(* Logix 5000 project; controller NWGG 1756-L72 rev 35.12; software revision 35.00; part 18 of 19 *)
(* tags used below, declared in another part *)
   Auto_Start_Treatment : BOOL;
   Belt : udt_Motor[16];
   Belts_Ready : BOOL;
   Bin_Gate_Test : BOOL;
   Bin_Open_test : BOOL;
   Bins_Rqd : BOOL;
   ckIDX : DINT;
   cntTransferTime : COUNTER;
   cntTreatTime : COUNTER;
   Concrete_Belts_Ready : BOOL;
   Concrete_Leg : udt_Motor;
   Current_Dist_List_IDX : DINT;
   Finish_Treat_Ok : BOOL;
   IDX : DINT;
   Loadout_Bin : udt_Loadout_Bin[29];
   Loadout_K_Valve : udt_Loadout_K_Valve[2];
   Longest_Treat_Stop_IDX : DINT;
   Loop_Idx : DINT;
   Manual_Mode : BOOL;
   Pause_Load_By_Time : BOOL[32];
   Pause_Load_By_Weight : BOOL[32];
   Pause_Load_Expired : DINT[2];
   Pause_Load_Pre : DINT[2];
   Pause_Transfer_By_Time : BOOL;
   Pause_Transfer_Load_Expired : DINT;
   Pause_Transfer_Msc : DINT;
   Pause_Transfer_Pre : DINT;
   Remote_Pause_Treat : BOOL;
   Reset_Remote_Pause : BOOL;
   Reset_Treat_Chemicals : BOOL;
   Reversing_Belt_Bypass_Valve : BOOL;
   Reversing_Belt_Reversed : BOOL;
   Start_Treat_Belts_Enabled : BOOL;
   Steel_Rqd_Belts_Running : BOOL;
   Stop_Treater : BOOL;
   Target_Weight : DINT[2];
   tmr_Pause_Load_Timer : TIMER[2];
   tmr_Pause_Transfer_Timer : TIMER;
   tmrBin_Delay_Start : TIMER[30];
   tmrDelayTreatStart : TIMER;
   tmrDelayTreatStop : TIMER;
   tmrResetChemicals : TIMER;
   tmrTransferTime : TIMER;
   tmrTreatTime : TIMER;
   Transfer_Batch_Status : DINT;
   Transfer_Belts_Starting : BOOL;
   Transfer_From_IDX : DINT;
   Transfer_Interlock : BOOL;
   Transfer_To_IDX : DINT;
   TransferHours : DINT;
   TransferMinuets : DINT;
   TransferSeconds : DINT;
   Treat_Batch_Status : DINT;
   Treat_Bin_Gates_Opened : BOOL;
   Treat_Bins_Open : BOOL;
   Treat_Interlock : BOOL;
   Treater_Loadout : udt_Treater_Loadout;
   TreatHours : DINT;
   Treatment_Running : BOOL;
   Treatment_Started : BOOL;
   TreatMinuets : DINT;
   TreatSeconds : DINT;
   Use_Concrete_Side_Treat : BOOL;
   Use_Steel_Side_Treat : BOOL;
   Use_Steel_Transfer_Bins : BOOL;
   tmrSetWaterOil : TIMER;
   Treater_Remote_Out : DINT;
   Truck_Scales : udt_Truck_Scale[2];
(* SeedLoadoutMain, continued *)

ROUTINE tmrTest   (* ladder *)
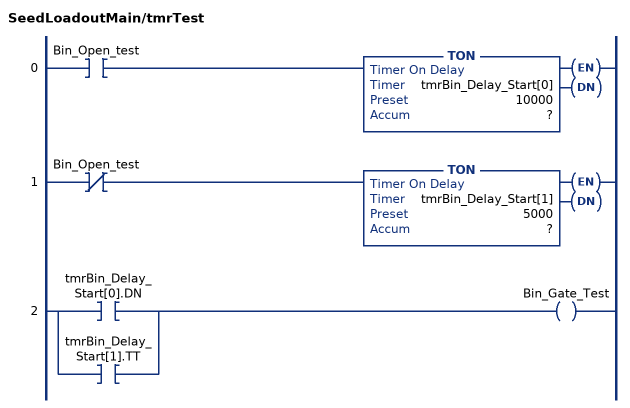
   0: XIC(Bin_Open_test)TON(tmrBin_Delay_Start[0],?,?);
   1: XIO(Bin_Open_test)TON(tmrBin_Delay_Start[1],?,?);
   2: [XIC(tmrBin_Delay_Start[0].DN) ,XIC(tmrBin_Delay_Start[1].TT) ]OTE(Bin_Gate_Test);
END_ROUTINE

ROUTINE Transfer_Belt_Batch_Ready   (* ladder *)
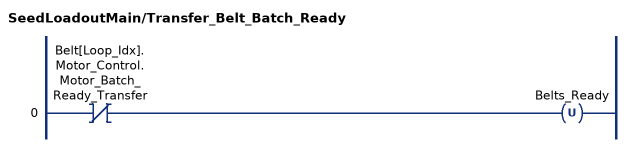
   0: XIO(Belt[Loop_Idx].Motor_Control.Motor_Batch_Ready_Transfer)OTU(Belts_Ready);
END_ROUTINE

ROUTINE Transfer_Belt_Start   (* ladder *)
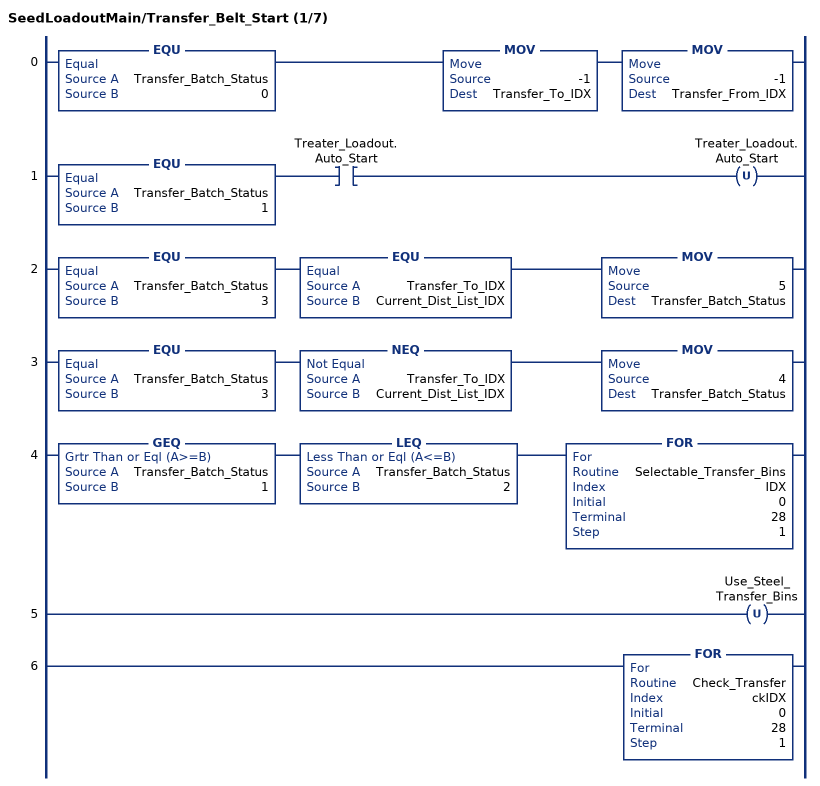
   0: EQU(Transfer_Batch_Status,0)MOV(-1,Transfer_To_IDX)MOV(-1,Transfer_From_IDX);
   1: EQU(Transfer_Batch_Status,1)XIC(Treater_Loadout.Auto_Start)OTU(Treater_Loadout.Auto_Start);
   2: EQU(Transfer_Batch_Status,3)EQU(Transfer_To_IDX,Current_Dist_List_IDX)MOV(5,Transfer_Batch_Status);
   3: EQU(Transfer_Batch_Status,3)NEQ(Transfer_To_IDX,Current_Dist_List_IDX)MOV(4,Transfer_Batch_Status);
   4: GEQ(Transfer_Batch_Status,1)LEQ(Transfer_Batch_Status,2)FOR(Selectable_Transfer_Bins,IDX,0,28,1);
   5: OTU(Use_Steel_Transfer_Bins);
   6: FOR(Check_Transfer,ckIDX,0,28,1);
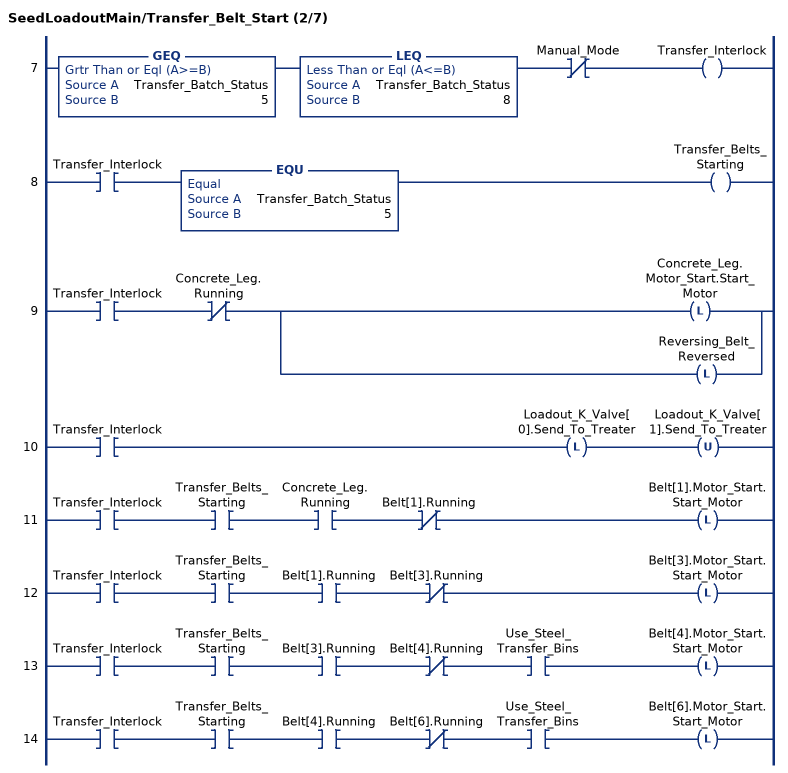
   7: GEQ(Transfer_Batch_Status,5)LEQ(Transfer_Batch_Status,8)XIO(Manual_Mode)OTE(Transfer_Interlock);
   8: XIC(Transfer_Interlock)EQU(Transfer_Batch_Status,5)OTE(Transfer_Belts_Starting);
   9: XIC(Transfer_Interlock)XIO(Concrete_Leg.Running)[OTL(Concrete_Leg.Motor_Start.Start_Motor) ,OTL(Reversing_Belt_Reversed) ];
   10: XIC(Transfer_Interlock)OTL(Loadout_K_Valve[0].Send_To_Treater)OTU(Loadout_K_Valve[1].Send_To_Treater);
   11: XIC(Transfer_Interlock)XIC(Transfer_Belts_Starting)XIC(Concrete_Leg.Running)XIO(Belt[1].Running)OTL(Belt[1].Motor_Start.Start_Motor);
   12: XIC(Transfer_Interlock)XIC(Transfer_Belts_Starting)XIC(Belt[1].Running)XIO(Belt[3].Running)OTL(Belt[3].Motor_Start.Start_Motor);
   13: XIC(Transfer_Interlock)XIC(Transfer_Belts_Starting)XIC(Belt[3].Running)XIO(Belt[4].Running)XIC(Use_Steel_Transfer_Bins)OTL(Belt[4].Motor_Start.Start_Motor);
   14: XIC(Transfer_Interlock)XIC(Transfer_Belts_Starting)XIC(Belt[4].Running)XIO(Belt[6].Running)XIC(Use_Steel_Transfer_Bins)OTL(Belt[6].Motor_Start.Start_Motor);
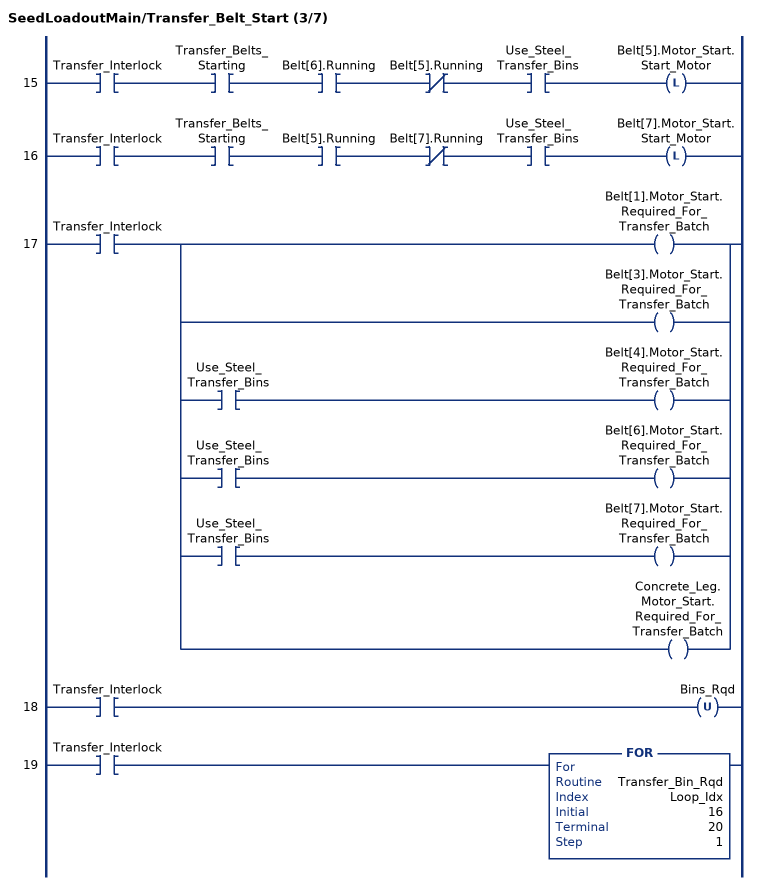
   15: XIC(Transfer_Interlock)XIC(Transfer_Belts_Starting)XIC(Belt[6].Running)XIO(Belt[5].Running)XIC(Use_Steel_Transfer_Bins)OTL(Belt[5].Motor_Start.Start_Motor);
   16: XIC(Transfer_Interlock)XIC(Transfer_Belts_Starting)XIC(Belt[5].Running)XIO(Belt[7].Running)XIC(Use_Steel_Transfer_Bins)OTL(Belt[7].Motor_Start.Start_Motor);
   17: XIC(Transfer_Interlock)[OTE(Belt[1].Motor_Start.Required_For_Transfer_Batch) ,OTE(Belt[3].Motor_Start.Required_For_Transfer_Batch) ,XIC(Use_Steel_Transfer_Bins) OTE(Belt[4].Motor_Start.Required_For_Transfer_Batch) ,XIC(Use_Steel_Transfer_Bins) OTE(Belt[6].Motor_Start.Required_For_Transfer_Batch) ,XIC(Use_Steel_Transfer_Bins) OTE(Belt[7].Motor_Start.Required_For_Transfer_Batch) ,OTE(Concrete_Leg.Motor_Start.Required_For_Transfer_Batch) ];
   18: XIC(Transfer_Interlock)OTU(Bins_Rqd);
   19: XIC(Transfer_Interlock)FOR(Transfer_Bin_Rqd,Loop_Idx,16,20,1);
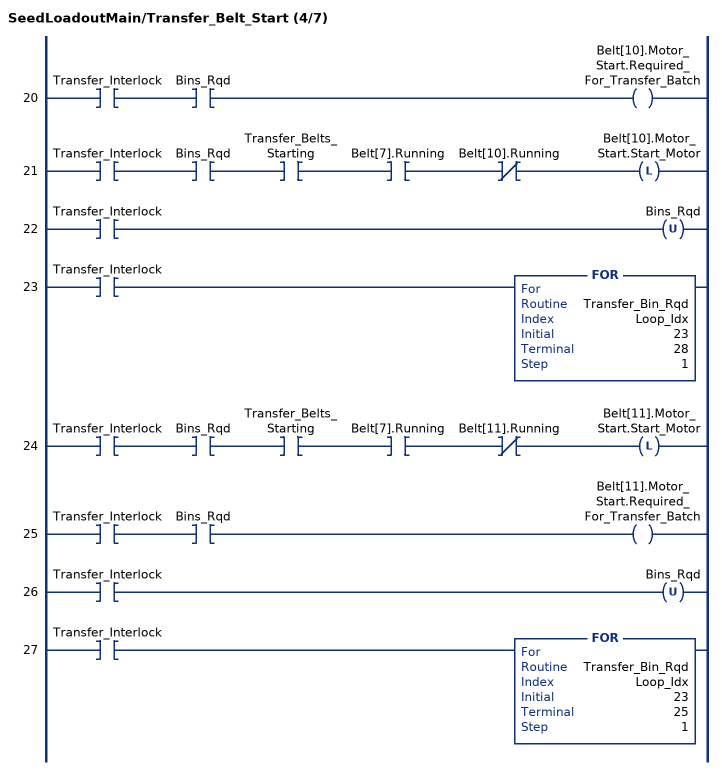
   20: XIC(Transfer_Interlock)XIC(Bins_Rqd)OTE(Belt[10].Motor_Start.Required_For_Transfer_Batch);
   21: XIC(Transfer_Interlock)XIC(Bins_Rqd)XIC(Transfer_Belts_Starting)XIC(Belt[7].Running)XIO(Belt[10].Running)OTL(Belt[10].Motor_Start.Start_Motor);
   22: XIC(Transfer_Interlock)OTU(Bins_Rqd);
   23: XIC(Transfer_Interlock)FOR(Transfer_Bin_Rqd,Loop_Idx,23,28,1);
   24: XIC(Transfer_Interlock)XIC(Bins_Rqd)XIC(Transfer_Belts_Starting)XIC(Belt[7].Running)XIO(Belt[11].Running)OTL(Belt[11].Motor_Start.Start_Motor);
   25: XIC(Transfer_Interlock)XIC(Bins_Rqd)OTE(Belt[11].Motor_Start.Required_For_Transfer_Batch);
   26: XIC(Transfer_Interlock)OTU(Bins_Rqd);
   27: XIC(Transfer_Interlock)FOR(Transfer_Bin_Rqd,Loop_Idx,23,25,1);
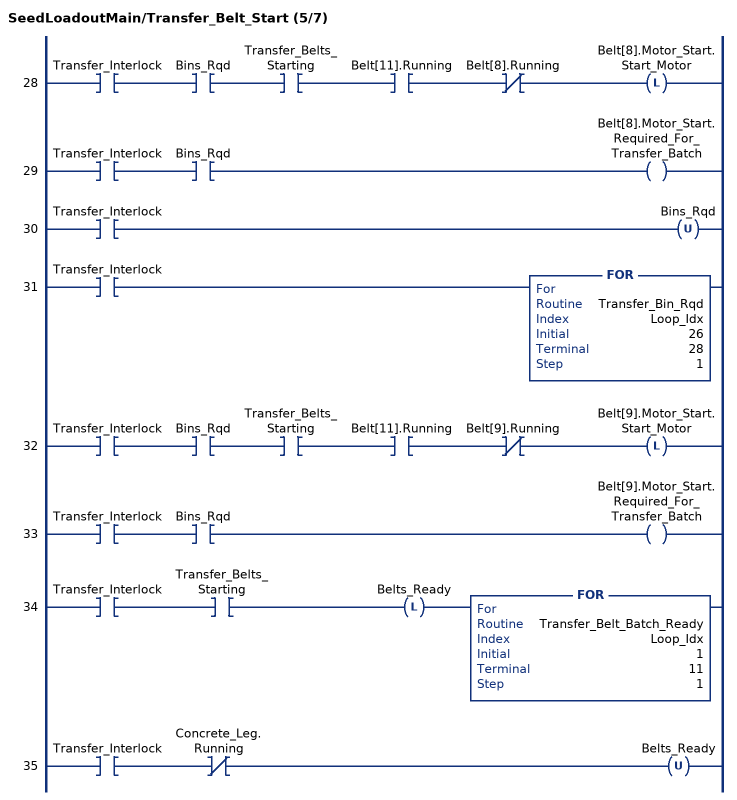
   28: XIC(Transfer_Interlock)XIC(Bins_Rqd)XIC(Transfer_Belts_Starting)XIC(Belt[11].Running)XIO(Belt[8].Running)OTL(Belt[8].Motor_Start.Start_Motor);
   29: XIC(Transfer_Interlock)XIC(Bins_Rqd)OTE(Belt[8].Motor_Start.Required_For_Transfer_Batch);
   30: XIC(Transfer_Interlock)OTU(Bins_Rqd);
   31: XIC(Transfer_Interlock)FOR(Transfer_Bin_Rqd,Loop_Idx,26,28,1);
   32: XIC(Transfer_Interlock)XIC(Bins_Rqd)XIC(Transfer_Belts_Starting)XIC(Belt[11].Running)XIO(Belt[9].Running)OTL(Belt[9].Motor_Start.Start_Motor);
   33: XIC(Transfer_Interlock)XIC(Bins_Rqd)OTE(Belt[9].Motor_Start.Required_For_Transfer_Batch);
   34: XIC(Transfer_Interlock)XIC(Transfer_Belts_Starting)OTL(Belts_Ready)FOR(Transfer_Belt_Batch_Ready,Loop_Idx,1,11,1);
   35: XIC(Transfer_Interlock)XIO(Concrete_Leg.Running)OTU(Belts_Ready);
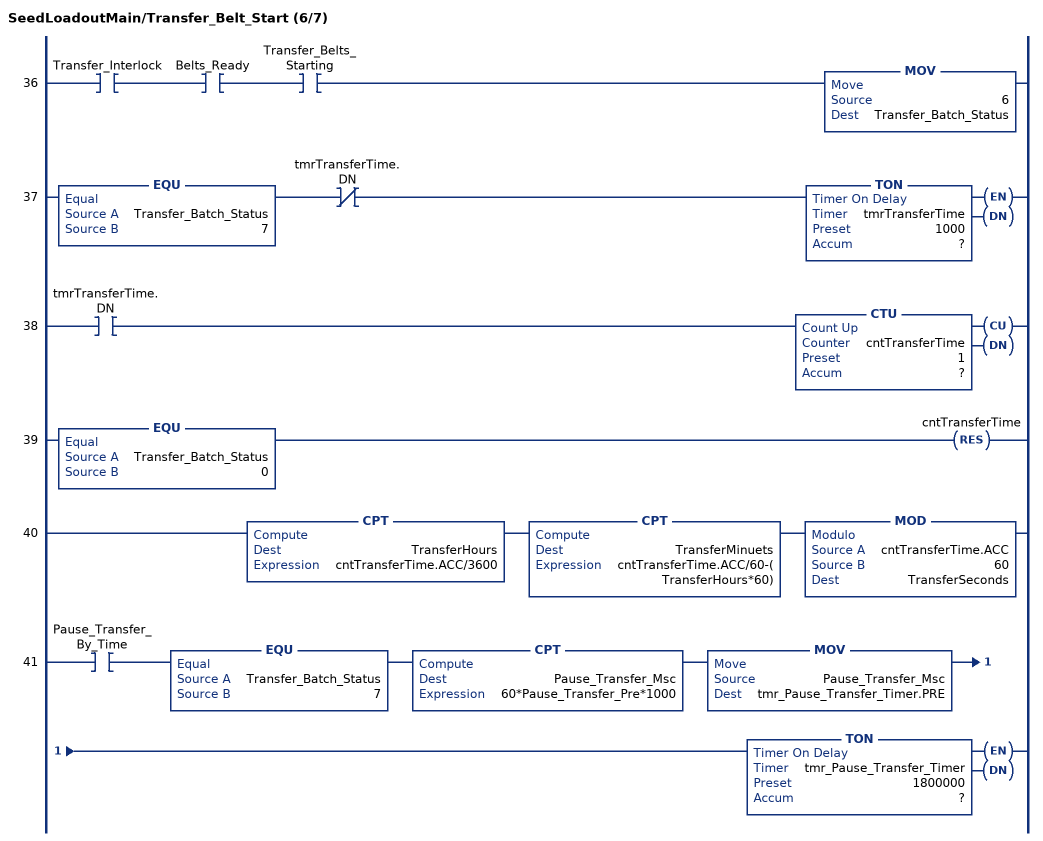
   36: XIC(Transfer_Interlock)XIC(Belts_Ready)XIC(Transfer_Belts_Starting)MOV(6,Transfer_Batch_Status);
   37: EQU(Transfer_Batch_Status,7)XIO(tmrTransferTime.DN)TON(tmrTransferTime,?,?);
   38: XIC(tmrTransferTime.DN)CTU(cntTransferTime,?,?);
   39: EQU(Transfer_Batch_Status,0)RES(cntTransferTime);
   40: CPT(TransferHours,cntTransferTime.ACC/3600)CPT(TransferMinuets,cntTransferTime.ACC/60-(TransferHours*60))MOD(cntTransferTime.ACC,60,TransferSeconds);
   41: XIC(Pause_Transfer_By_Time)EQU(Transfer_Batch_Status,7)CPT(Pause_Transfer_Msc,60*Pause_Transfer_Pre*1000)MOV(Pause_Transfer_Msc,tmr_Pause_Transfer_Timer.PRE)TON(tmr_Pause_Transfer_Timer,?,?);
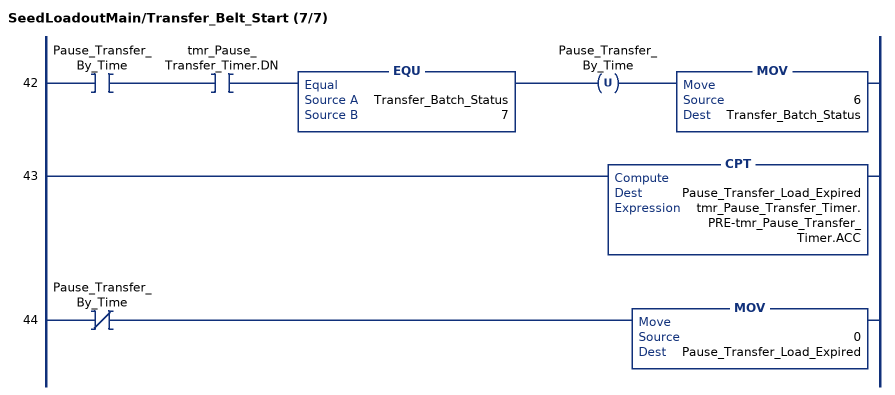
   42: XIC(Pause_Transfer_By_Time)XIC(tmr_Pause_Transfer_Timer.DN)EQU(Transfer_Batch_Status,7)OTU(Pause_Transfer_By_Time)MOV(6,Transfer_Batch_Status);
   43: CPT(Pause_Transfer_Load_Expired,tmr_Pause_Transfer_Timer.PRE-tmr_Pause_Transfer_Timer.ACC);
   44: XIO(Pause_Transfer_By_Time)MOV(0,Pause_Transfer_Load_Expired);
END_ROUTINE

ROUTINE Transfer_Bin_Rqd   (* ladder *)
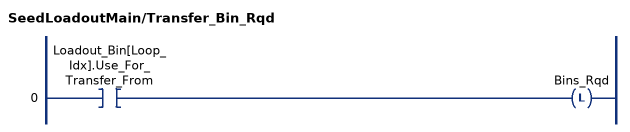
   0: XIC(Loadout_Bin[Loop_Idx].Use_For_Transfer_From)OTL(Bins_Rqd);
END_ROUTINE

ROUTINE Treat_Belt_Batch_Ready   (* ladder *)
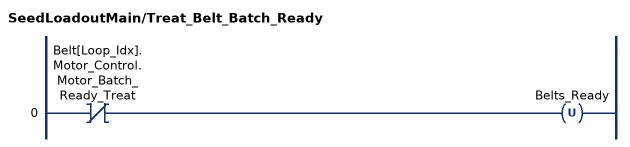
   0: XIO(Belt[Loop_Idx].Motor_Control.Motor_Batch_Ready_Treat)OTU(Belts_Ready);
END_ROUTINE

ROUTINE Treat_Belt_Start   (* ladder *)
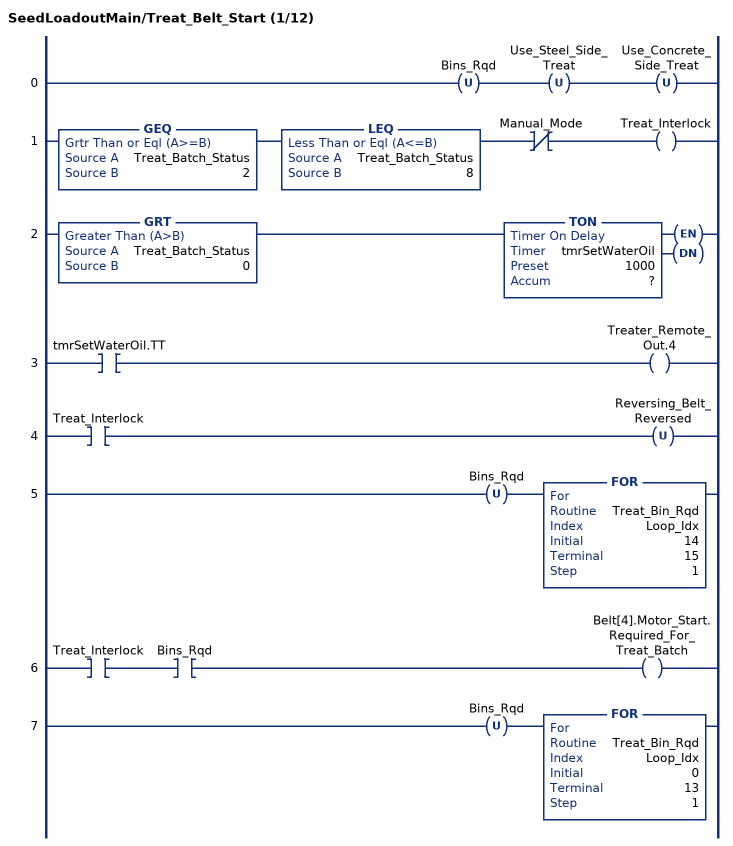
   0: OTU(Bins_Rqd)OTU(Use_Steel_Side_Treat)OTU(Use_Concrete_Side_Treat);
   1: GEQ(Treat_Batch_Status,2)LEQ(Treat_Batch_Status,8)XIO(Manual_Mode)OTE(Treat_Interlock);
   2: GRT(Treat_Batch_Status,0)TON(tmrSetWaterOil,?,?);
   3: XIC(tmrSetWaterOil.TT)OTE(Treater_Remote_Out.4);
   4: XIC(Treat_Interlock)OTU(Reversing_Belt_Reversed);
   5: OTU(Bins_Rqd)FOR(Treat_Bin_Rqd,Loop_Idx,14,15,1);
   6: XIC(Treat_Interlock)XIC(Bins_Rqd)OTE(Belt[4].Motor_Start.Required_For_Treat_Batch);
   7: OTU(Bins_Rqd)FOR(Treat_Bin_Rqd,Loop_Idx,0,13,1);
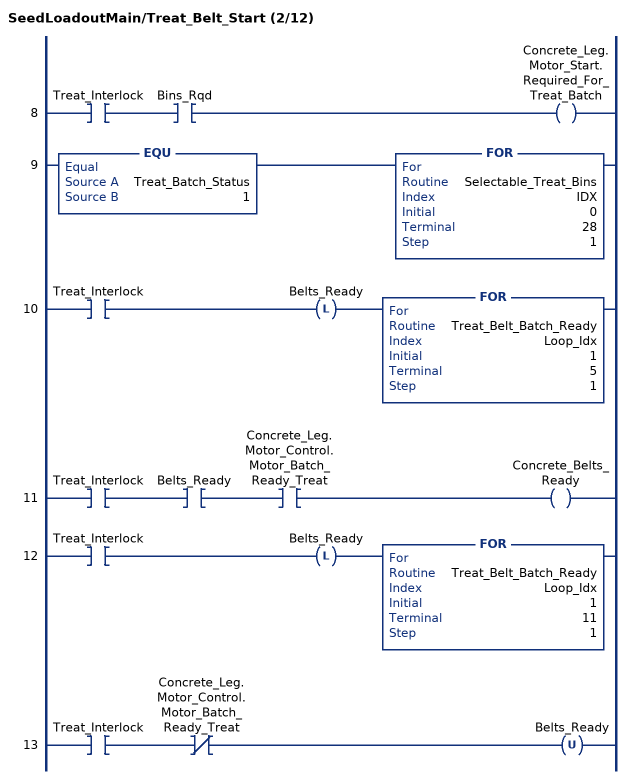
   8: XIC(Treat_Interlock)XIC(Bins_Rqd)OTE(Concrete_Leg.Motor_Start.Required_For_Treat_Batch);
   9: EQU(Treat_Batch_Status,1)FOR(Selectable_Treat_Bins,IDX,0,28,1);
   10: XIC(Treat_Interlock)OTL(Belts_Ready)FOR(Treat_Belt_Batch_Ready,Loop_Idx,1,5,1);
   11: XIC(Treat_Interlock)XIC(Belts_Ready)XIC(Concrete_Leg.Motor_Control.Motor_Batch_Ready_Treat)OTE(Concrete_Belts_Ready);
   12: XIC(Treat_Interlock)OTL(Belts_Ready)FOR(Treat_Belt_Batch_Ready,Loop_Idx,1,11,1);
   13: XIC(Treat_Interlock)XIO(Concrete_Leg.Motor_Control.Motor_Batch_Ready_Treat)OTU(Belts_Ready);
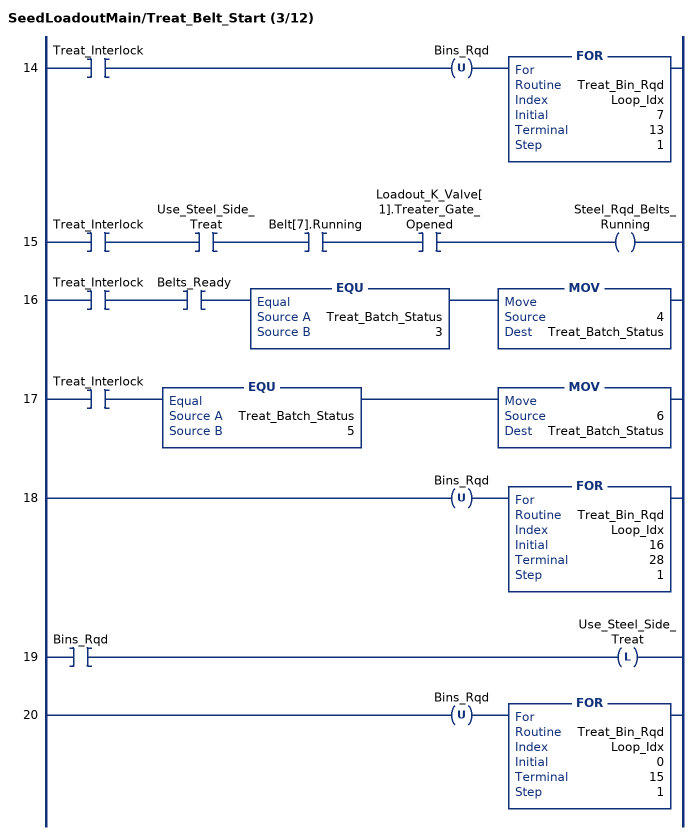
   14: XIC(Treat_Interlock)OTU(Bins_Rqd)FOR(Treat_Bin_Rqd,Loop_Idx,7,13,1);
   15: XIC(Treat_Interlock)XIC(Use_Steel_Side_Treat)XIC(Belt[7].Running)XIC(Loadout_K_Valve[1].Treater_Gate_Opened)OTE(Steel_Rqd_Belts_Running);
   16: XIC(Treat_Interlock)XIC(Belts_Ready)EQU(Treat_Batch_Status,3)MOV(4,Treat_Batch_Status);
   17: XIC(Treat_Interlock)EQU(Treat_Batch_Status,5)MOV(6,Treat_Batch_Status);
   18: OTU(Bins_Rqd)FOR(Treat_Bin_Rqd,Loop_Idx,16,28,1);
   19: XIC(Bins_Rqd)OTL(Use_Steel_Side_Treat);
   20: OTU(Bins_Rqd)FOR(Treat_Bin_Rqd,Loop_Idx,0,15,1);
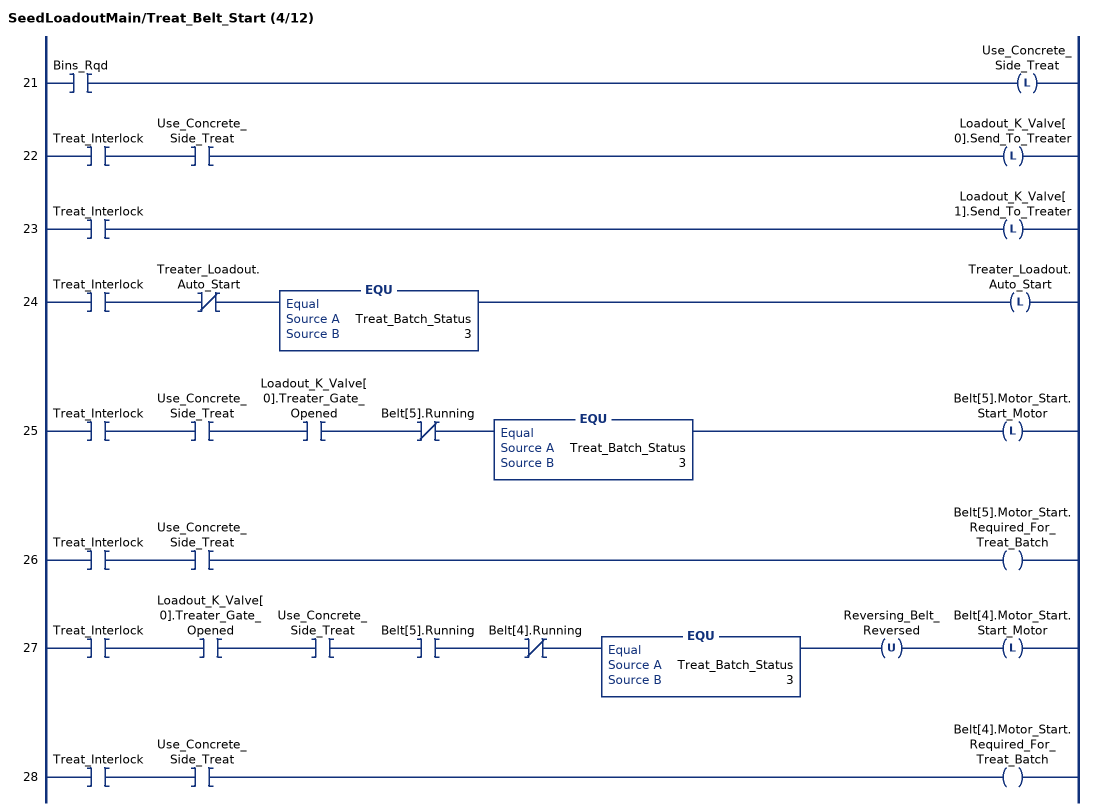
   21: XIC(Bins_Rqd)OTL(Use_Concrete_Side_Treat);
   22: XIC(Treat_Interlock)XIC(Use_Concrete_Side_Treat)OTL(Loadout_K_Valve[0].Send_To_Treater);
   23: XIC(Treat_Interlock)OTL(Loadout_K_Valve[1].Send_To_Treater);
   24: XIC(Treat_Interlock)XIO(Treater_Loadout.Auto_Start)EQU(Treat_Batch_Status,3)OTL(Treater_Loadout.Auto_Start);
   25: XIC(Treat_Interlock)XIC(Use_Concrete_Side_Treat)XIC(Loadout_K_Valve[0].Treater_Gate_Opened)XIO(Belt[5].Running)EQU(Treat_Batch_Status,3)OTL(Belt[5].Motor_Start.Start_Motor);
   26: XIC(Treat_Interlock)XIC(Use_Concrete_Side_Treat)OTE(Belt[5].Motor_Start.Required_For_Treat_Batch);
   27: XIC(Treat_Interlock)XIC(Loadout_K_Valve[0].Treater_Gate_Opened)XIC(Use_Concrete_Side_Treat)XIC(Belt[5].Running)XIO(Belt[4].Running)EQU(Treat_Batch_Status,3)OTU(Reversing_Belt_Reversed)OTL(Belt[4].Motor_Start.Start_Motor);
   28: XIC(Treat_Interlock)XIC(Use_Concrete_Side_Treat)OTE(Belt[4].Motor_Start.Required_For_Treat_Batch);
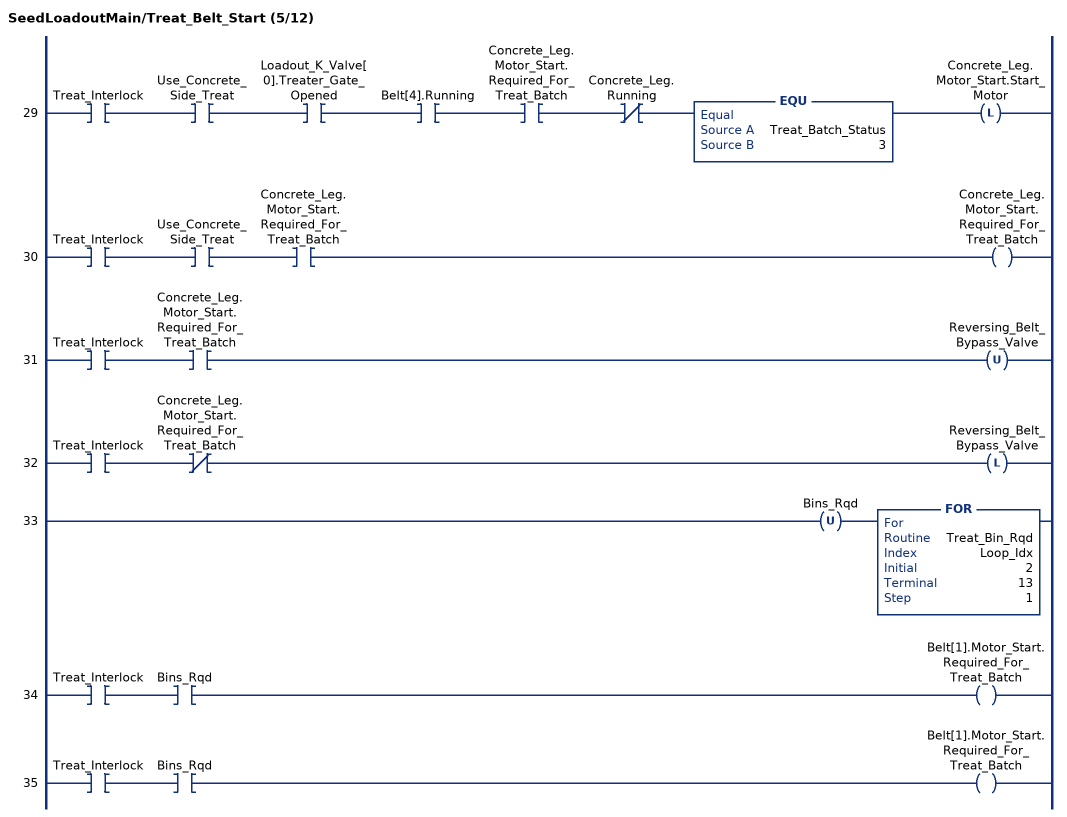
   29: XIC(Treat_Interlock)XIC(Use_Concrete_Side_Treat)XIC(Loadout_K_Valve[0].Treater_Gate_Opened)XIC(Belt[4].Running)XIC(Concrete_Leg.Motor_Start.Required_For_Treat_Batch)XIO(Concrete_Leg.Running)EQU(Treat_Batch_Status,3)OTL(Concrete_Leg.Motor_Start.Start_Motor);
   30: XIC(Treat_Interlock)XIC(Use_Concrete_Side_Treat)XIC(Concrete_Leg.Motor_Start.Required_For_Treat_Batch)OTE(Concrete_Leg.Motor_Start.Required_For_Treat_Batch);
   31: XIC(Treat_Interlock)XIC(Concrete_Leg.Motor_Start.Required_For_Treat_Batch)OTU(Reversing_Belt_Bypass_Valve);
   32: XIC(Treat_Interlock)XIO(Concrete_Leg.Motor_Start.Required_For_Treat_Batch)OTL(Reversing_Belt_Bypass_Valve);
   33: OTU(Bins_Rqd)FOR(Treat_Bin_Rqd,Loop_Idx,2,13,1);
   34: XIC(Treat_Interlock)XIC(Bins_Rqd)OTE(Belt[1].Motor_Start.Required_For_Treat_Batch);
   35: XIC(Treat_Interlock)XIC(Bins_Rqd)OTE(Belt[1].Motor_Start.Required_For_Treat_Batch);
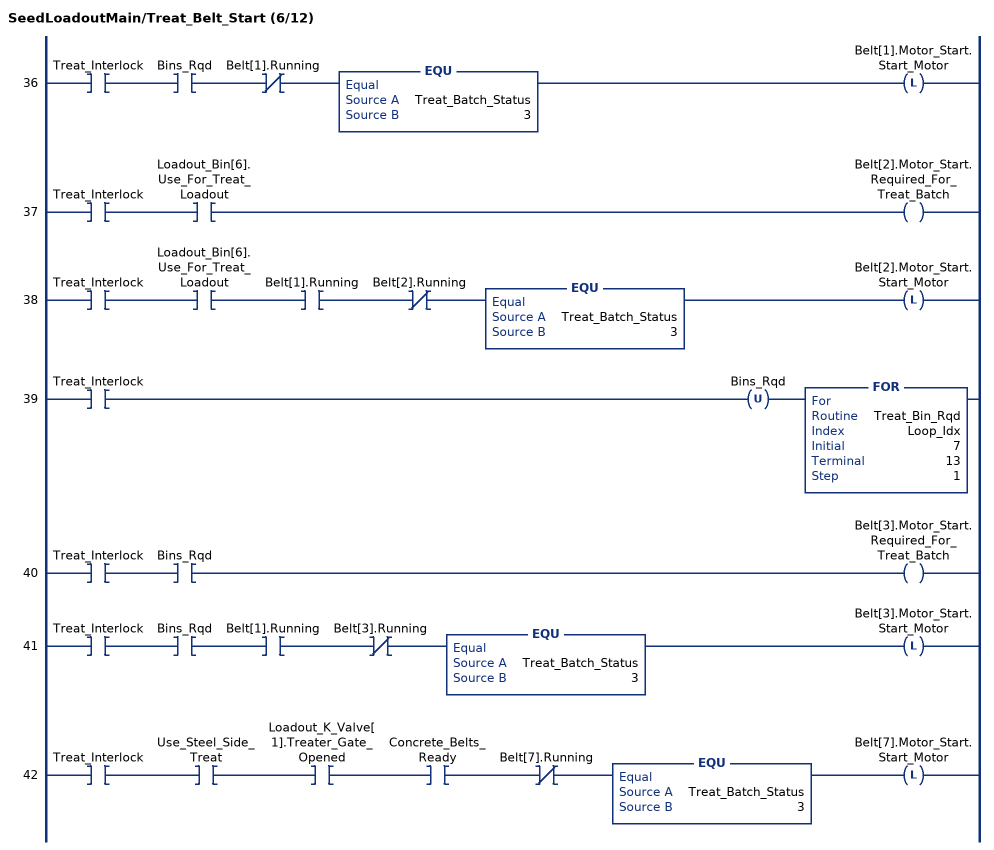
   36: XIC(Treat_Interlock)XIC(Bins_Rqd)XIO(Belt[1].Running)EQU(Treat_Batch_Status,3)OTL(Belt[1].Motor_Start.Start_Motor);
   37: XIC(Treat_Interlock)XIC(Loadout_Bin[6].Use_For_Treat_Loadout)OTE(Belt[2].Motor_Start.Required_For_Treat_Batch);
   38: XIC(Treat_Interlock)XIC(Loadout_Bin[6].Use_For_Treat_Loadout)XIC(Belt[1].Running)XIO(Belt[2].Running)EQU(Treat_Batch_Status,3)OTL(Belt[2].Motor_Start.Start_Motor);
   39: XIC(Treat_Interlock)OTU(Bins_Rqd)FOR(Treat_Bin_Rqd,Loop_Idx,7,13,1);
   40: XIC(Treat_Interlock)XIC(Bins_Rqd)OTE(Belt[3].Motor_Start.Required_For_Treat_Batch);
   41: XIC(Treat_Interlock)XIC(Bins_Rqd)XIC(Belt[1].Running)XIO(Belt[3].Running)EQU(Treat_Batch_Status,3)OTL(Belt[3].Motor_Start.Start_Motor);
   42: XIC(Treat_Interlock)XIC(Use_Steel_Side_Treat)XIC(Loadout_K_Valve[1].Treater_Gate_Opened)XIC(Concrete_Belts_Ready)XIO(Belt[7].Running)EQU(Treat_Batch_Status,3)OTL(Belt[7].Motor_Start.Start_Motor);
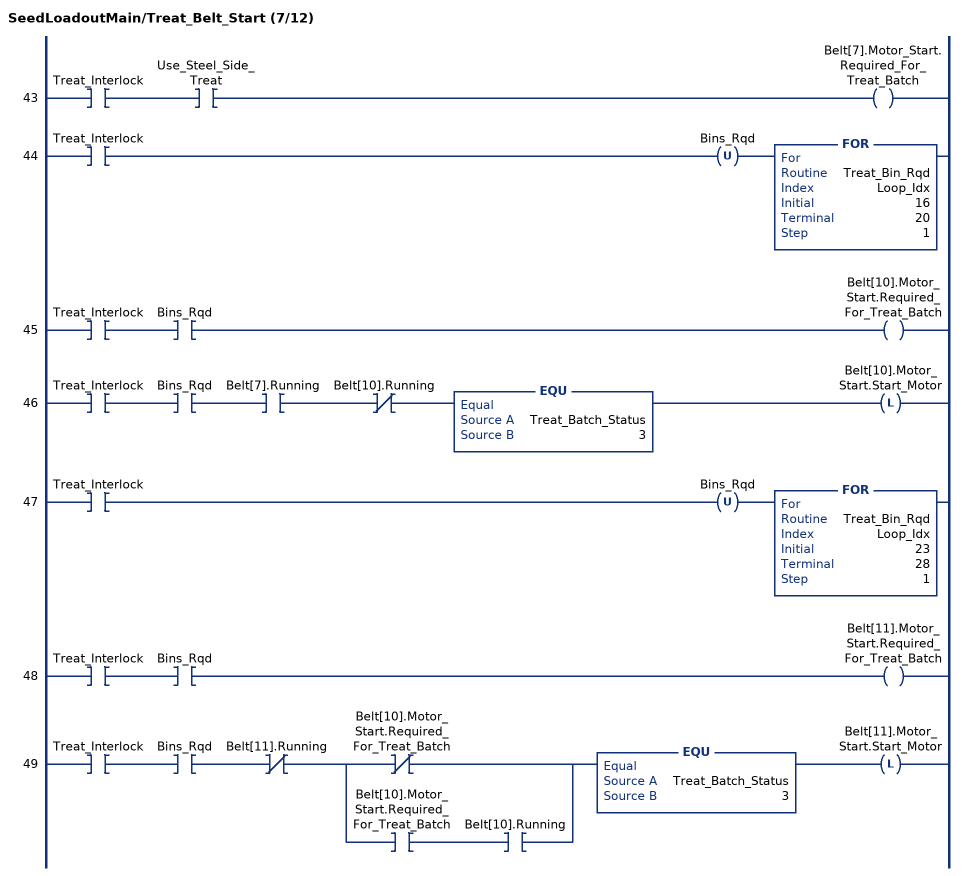
   43: XIC(Treat_Interlock)XIC(Use_Steel_Side_Treat)OTE(Belt[7].Motor_Start.Required_For_Treat_Batch);
   44: XIC(Treat_Interlock)OTU(Bins_Rqd)FOR(Treat_Bin_Rqd,Loop_Idx,16,20,1);
   45: XIC(Treat_Interlock)XIC(Bins_Rqd)OTE(Belt[10].Motor_Start.Required_For_Treat_Batch);
   46: XIC(Treat_Interlock)XIC(Bins_Rqd)XIC(Belt[7].Running)XIO(Belt[10].Running)EQU(Treat_Batch_Status,3)OTL(Belt[10].Motor_Start.Start_Motor);
   47: XIC(Treat_Interlock)OTU(Bins_Rqd)FOR(Treat_Bin_Rqd,Loop_Idx,23,28,1);
   48: XIC(Treat_Interlock)XIC(Bins_Rqd)OTE(Belt[11].Motor_Start.Required_For_Treat_Batch);
   49: XIC(Treat_Interlock)XIC(Bins_Rqd)XIO(Belt[11].Running)[XIO(Belt[10].Motor_Start.Required_For_Treat_Batch) ,XIC(Belt[10].Motor_Start.Required_For_Treat_Batch) XIC(Belt[10].Running) ]EQU(Treat_Batch_Status,3)OTL(Belt[11].Motor_Start.Start_Motor);
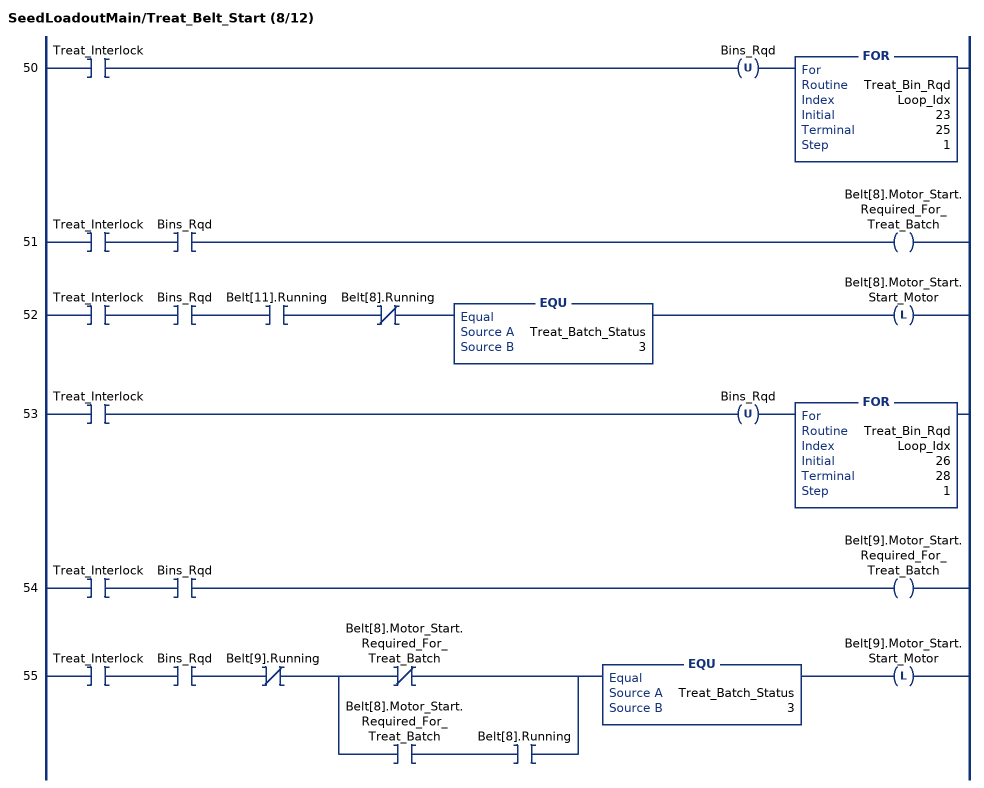
   50: XIC(Treat_Interlock)OTU(Bins_Rqd)FOR(Treat_Bin_Rqd,Loop_Idx,23,25,1);
   51: XIC(Treat_Interlock)XIC(Bins_Rqd)OTE(Belt[8].Motor_Start.Required_For_Treat_Batch);
   52: XIC(Treat_Interlock)XIC(Bins_Rqd)XIC(Belt[11].Running)XIO(Belt[8].Running)EQU(Treat_Batch_Status,3)OTL(Belt[8].Motor_Start.Start_Motor);
   53: XIC(Treat_Interlock)OTU(Bins_Rqd)FOR(Treat_Bin_Rqd,Loop_Idx,26,28,1);
   54: XIC(Treat_Interlock)XIC(Bins_Rqd)OTE(Belt[9].Motor_Start.Required_For_Treat_Batch);
   55: XIC(Treat_Interlock)XIC(Bins_Rqd)XIO(Belt[9].Running)[XIO(Belt[8].Motor_Start.Required_For_Treat_Batch) ,XIC(Belt[8].Motor_Start.Required_For_Treat_Batch) XIC(Belt[8].Running) ]EQU(Treat_Batch_Status,3)OTL(Belt[9].Motor_Start.Start_Motor);
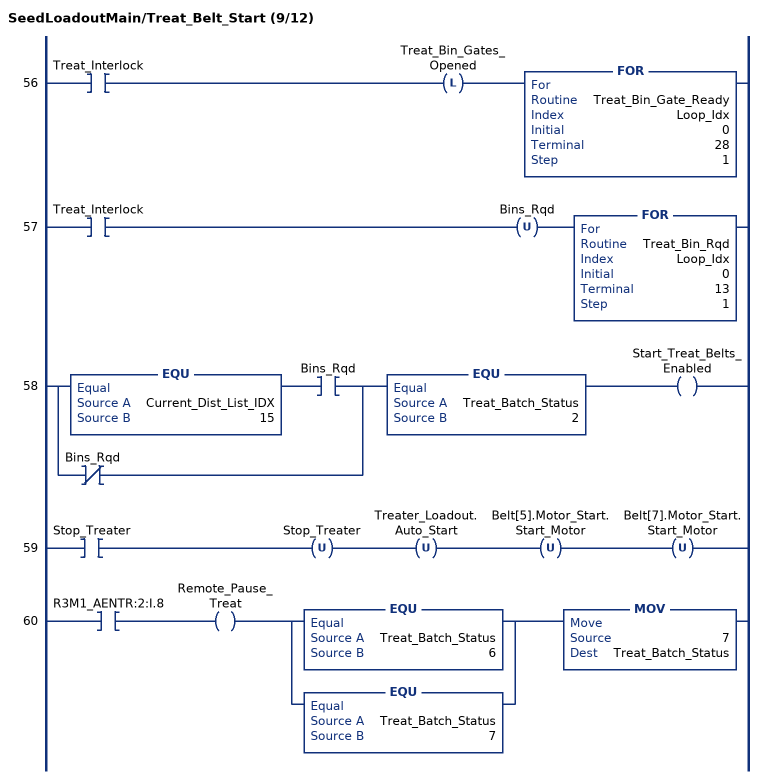
   56: XIC(Treat_Interlock)OTL(Treat_Bin_Gates_Opened)FOR(Treat_Bin_Gate_Ready,Loop_Idx,0,28,1);
   57: XIC(Treat_Interlock)OTU(Bins_Rqd)FOR(Treat_Bin_Rqd,Loop_Idx,0,13,1);
   58: [EQU(Current_Dist_List_IDX,15) XIC(Bins_Rqd) ,XIO(Bins_Rqd) ]EQU(Treat_Batch_Status,2)OTE(Start_Treat_Belts_Enabled);
   59: XIC(Stop_Treater)OTU(Stop_Treater)OTU(Treater_Loadout.Auto_Start)OTU(Belt[5].Motor_Start.Start_Motor)OTU(Belt[7].Motor_Start.Start_Motor);
   60: XIC(R3M1_AENTR:2:I.8)OTE(Remote_Pause_Treat)[EQU(Treat_Batch_Status,6) ,EQU(Treat_Batch_Status,7) ]MOV(7,Treat_Batch_Status);
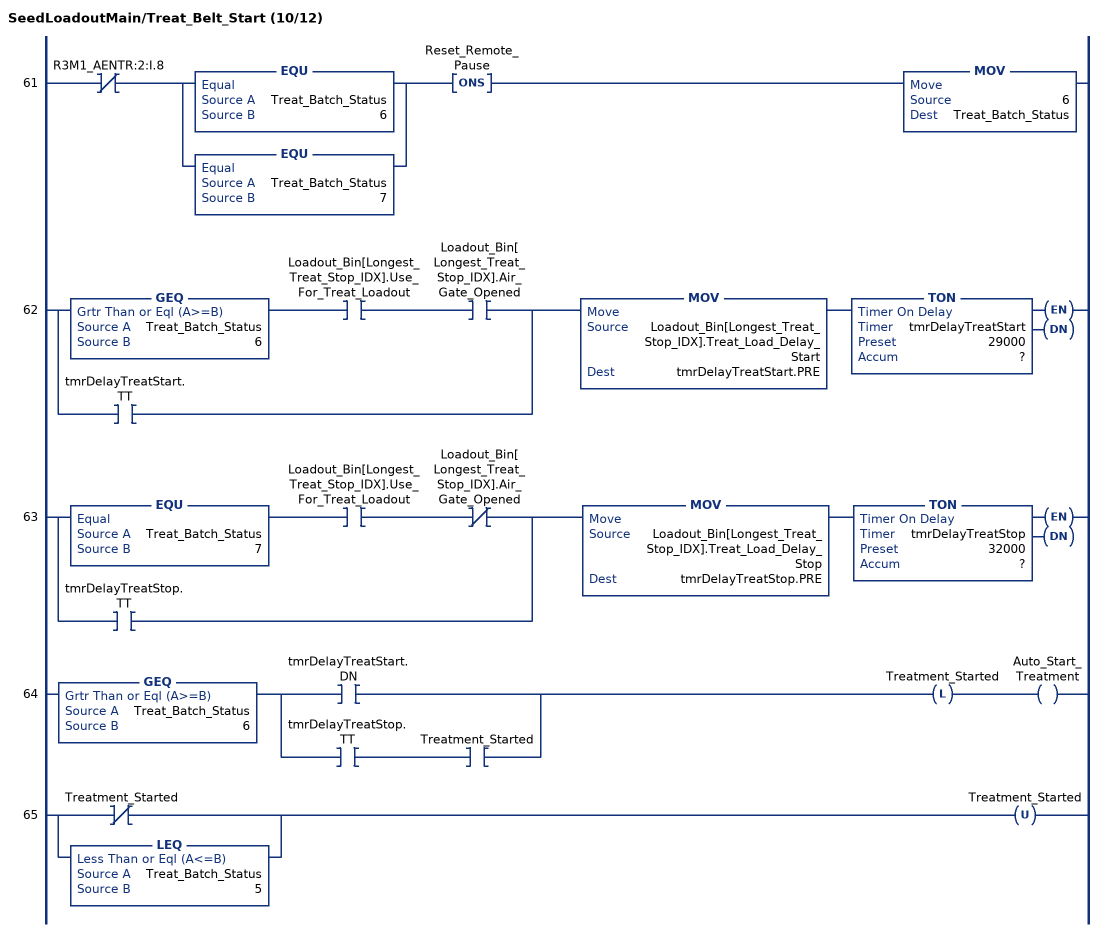
   61: XIO(R3M1_AENTR:2:I.8)[EQU(Treat_Batch_Status,6) ,EQU(Treat_Batch_Status,7) ]ONS(Reset_Remote_Pause)MOV(6,Treat_Batch_Status);
   62: [GEQ(Treat_Batch_Status,6) XIC(Loadout_Bin[Longest_Treat_Stop_IDX].Use_For_Treat_Loadout) XIC(Loadout_Bin[Longest_Treat_Stop_IDX].Air_Gate_Opened) ,XIC(tmrDelayTreatStart.TT) ]MOV(Loadout_Bin[Longest_Treat_Stop_IDX].Treat_Load_Delay_Start,tmrDelayTreatStart.PRE)TON(tmrDelayTreatStart,?,?);
   63: [EQU(Treat_Batch_Status,7) XIC(Loadout_Bin[Longest_Treat_Stop_IDX].Use_For_Treat_Loadout) XIO(Loadout_Bin[Longest_Treat_Stop_IDX].Air_Gate_Opened) ,XIC(tmrDelayTreatStop.TT) ]MOV(Loadout_Bin[Longest_Treat_Stop_IDX].Treat_Load_Delay_Stop,tmrDelayTreatStop.PRE)TON(tmrDelayTreatStop,?,?);
   64: GEQ(Treat_Batch_Status,6)[XIC(tmrDelayTreatStart.DN) ,XIC(tmrDelayTreatStop.TT) XIC(Treatment_Started) ]OTL(Treatment_Started)OTE(Auto_Start_Treatment);
   65: [XIO(Treatment_Started) ,LEQ(Treat_Batch_Status,5) ]OTU(Treatment_Started);
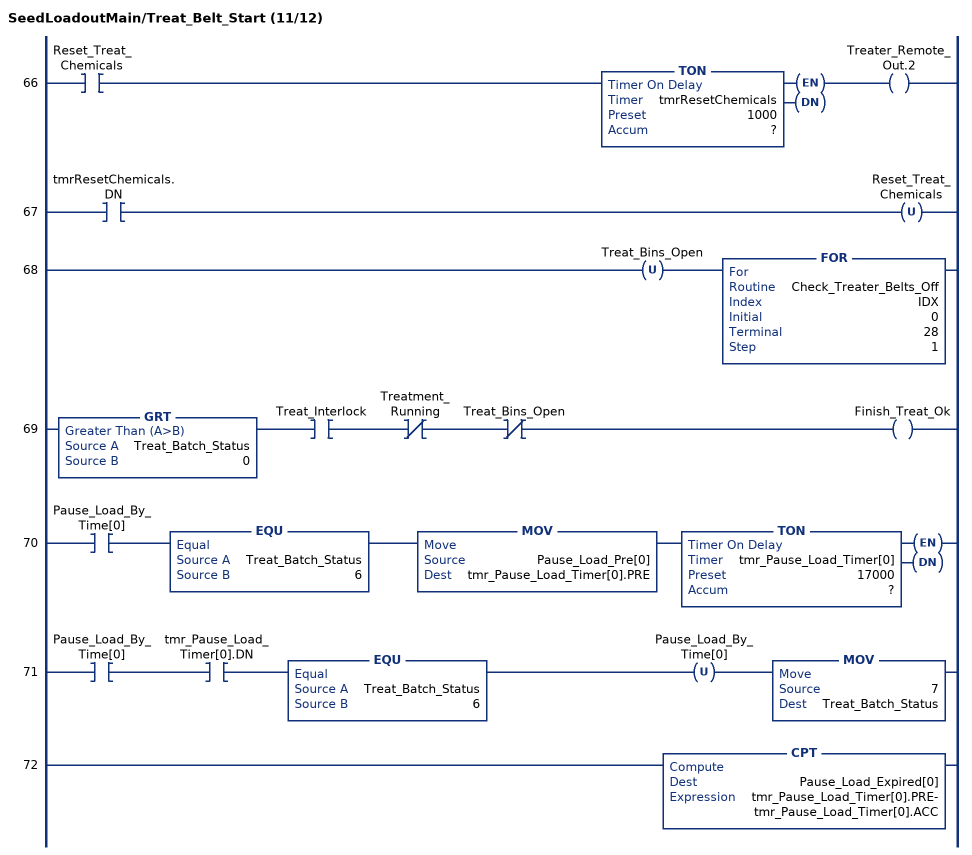
   66: XIC(Reset_Treat_Chemicals)TON(tmrResetChemicals,?,?)OTE(Treater_Remote_Out.2);
   67: XIC(tmrResetChemicals.DN)OTU(Reset_Treat_Chemicals);
   68: OTU(Treat_Bins_Open)FOR(Check_Treater_Belts_Off,IDX,0,28,1);
   69: GRT(Treat_Batch_Status,0)XIC(Treat_Interlock)XIO(Treatment_Running)XIO(Treat_Bins_Open)OTE(Finish_Treat_Ok);
   70: XIC(Pause_Load_By_Time[0])EQU(Treat_Batch_Status,6)MOV(Pause_Load_Pre[0],tmr_Pause_Load_Timer[0].PRE)TON(tmr_Pause_Load_Timer[0],?,?);
   71: XIC(Pause_Load_By_Time[0])XIC(tmr_Pause_Load_Timer[0].DN)EQU(Treat_Batch_Status,6)OTU(Pause_Load_By_Time[0])MOV(7,Treat_Batch_Status);
   72: CPT(Pause_Load_Expired[0],tmr_Pause_Load_Timer[0].PRE-tmr_Pause_Load_Timer[0].ACC);
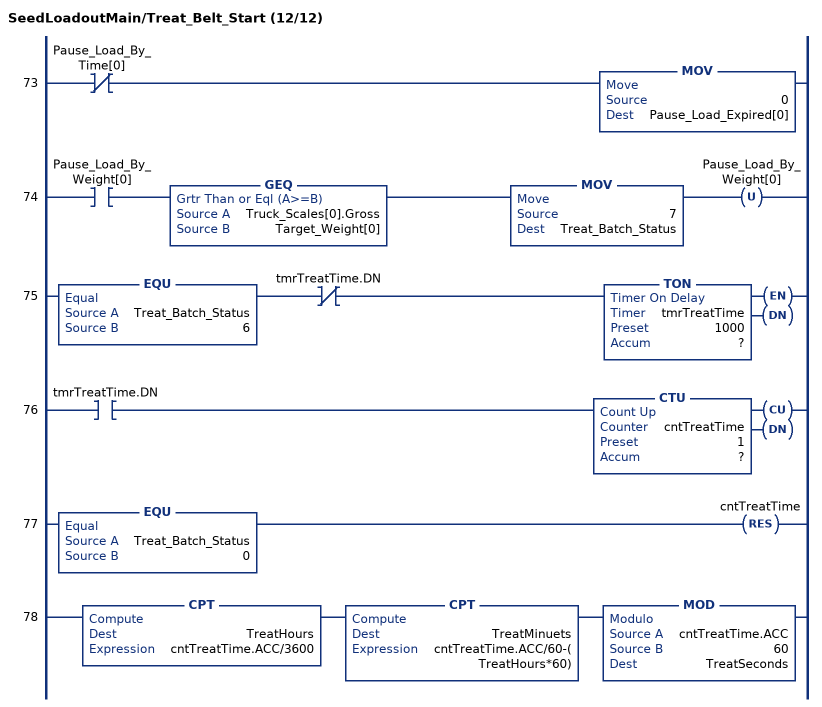
   73: XIO(Pause_Load_By_Time[0])MOV(0,Pause_Load_Expired[0]);
   74: XIC(Pause_Load_By_Weight[0])GEQ(Truck_Scales[0].Gross,Target_Weight[0])MOV(7,Treat_Batch_Status)OTU(Pause_Load_By_Weight[0]);
   75: EQU(Treat_Batch_Status,6)XIO(tmrTreatTime.DN)TON(tmrTreatTime,?,?);
   76: XIC(tmrTreatTime.DN)CTU(cntTreatTime,?,?);
   77: EQU(Treat_Batch_Status,0)RES(cntTreatTime);
   78: CPT(TreatHours,cntTreatTime.ACC/3600)CPT(TreatMinuets,cntTreatTime.ACC/60-(TreatHours*60))MOD(cntTreatTime.ACC,60,TreatSeconds);
END_ROUTINE
